(* IEC 61131-3 sources: University/4015/10 Feb 2026/LO2 LO3 - Mr Akbar/Programs/05 Precise Jog Pulse/build, 2 files *)

(* ---- plc.st ---- *)
TYPE
  LOGLEVEL : (CRITICAL, WARNING, INFO, DEBUG) := INFO;
END_TYPE

FUNCTION_BLOCK LOGGER
  VAR_INPUT
    TRIG : BOOL;
    MSG : STRING;
    LEVEL : LOGLEVEL := INFO;
  END_VAR
  VAR
    TRIG0 : BOOL;
  END_VAR

  IF TRIG AND NOT TRIG0 THEN
  {{
   LogMessage(GetFbVar(LEVEL),(char*)GetFbVar(MSG, .body),GetFbVar(MSG, .len));
  }}
  END_IF;
  TRIG0:=TRIG;
END_FUNCTION_BLOCK

PROGRAM program0
  VAR
    JOG_EDGE : BOOL;
    JOG_PULSE : BOOL;
  END_VAR
  VAR
    Duration : TIME := t#300ms;
    TP0 : TP;
    R_TRIG1 : R_TRIG;
  END_VAR

  R_TRIG1(CLK := JOG_EDGE);
  TP0(IN := R_TRIG1.Q, PT := Duration);
  JOG_PULSE := TP0.Q;
END_PROGRAM

CONFIGURATION Config0

  RESOURCE Res0 ON PLC
    TASK task0(INTERVAL := T#20ms,PRIORITY := 0);
    PROGRAM instance0 WITH task0 : program0;
  END_RESOURCE
END_CONFIGURATION

(* ---- generated_plc.st ---- *)
PROGRAM program0
  VAR
    JOG_EDGE AT %IX0.0 : BOOL;
    JOG_PULSE AT %M0.5 : BOOL;
  END_VAR
  VAR
    Duration : TIME := t#300ms;
    TP0 : TP;
    R_TRIG1 : R_TRIG;
  END_VAR

  R_TRIG1(CLK := JOG_EDGE);
  TP0(IN := R_TRIG1.Q, PT := Duration);
  JOG_PULSE := TP0.Q;
END_PROGRAM

CONFIGURATION Config0

  RESOURCE Res0 ON PLC
    TASK task0(INTERVAL := T#20ms,PRIORITY := 0);
    PROGRAM instance0 WITH task0 : program0;
  END_RESOURCE
END_CONFIGURATION
